Fanuc KAREL source: kt00298.KL

-- PROVISIONAL review KL for V770-1; original PC SHA256 92522de8097242ac7d6fa85fb294c7b0889a8dfae95d8bf3571cb3d213de84da
-- Incomplete behavior may be omitted. Consult companion uncertainty JSON. Do not deploy.
PROGRAM KT00298
%NOLOCKGROUP
VAR
  R1 : REAL
  R2 : REAL
  OUT : BOOLEAN
BEGIN
  -- UNRESOLVED_PC offsets 5-16; opcodes 2E,23
  -- UNRESOLVED_PC offsets 21-32; opcodes 2E,23
  -- UNRESOLVED_PC offsets 37-48; opcodes 2E,23
  -- UNRESOLVED_PC offsets 53-64; opcodes 2E,23
  -- UNRESOLVED_PC offsets 69-88; opcodes 21,21,6E,23
  -- UNRESOLVED_PC offsets 93-97; opcodes 7F
END KT00298
